// TwinCAT 3 PLC project AdsGo_Det
// Title: AdsClient_DeterministicTester
// Description: This project provides a series of programs and symbols to allow integration testing of ADS clients by utilising deterministic outputs on symbols based on writeable inputs (such as nSeed).
// ProgramVersion: 3.1.4026.25
// libraries:
//   Tc2_Standard, * (Beckhoff Automation GmbH)
//   Tc2_System, * (Beckhoff Automation GmbH)
//   Tc3_Module, * (Beckhoff Automation GmbH)
// project tree:
//   Lib/Arrays/ E_ArrayEnum.TcDUT, FB_ArrayTest.TcPOU, ST_Array.TcDUT, ST_ArrayBits.TcDUT
//   Lib/Attributes/ FB_AttributeTest.TcPOU
//   Lib/BitPacking/ FB_BitPackingTest.TcPOU, ST_BitPacking.TcDUT
//   Lib/Enums/ E_Int.TcDUT, E_Sparse.TcDUT, E_UInt.TcDUT, E_Default.TcDUT, E_Dint.TcDUT, E_Byte.TcDUT, E_Sint.TcDUT, E_USint.TcDUT, E_Word.TcDUT, E_ULint.TcDUT, E_UDint.TcDUT, E_Lint.TcDUT, E_DWord.TcDUT, E_LWord.TcDUT, E_Negative.TcDUT, FB_EnumTest.TcPOU
//   Lib/ FB_TickCounter.TcPOU
//   Lib/Gvl/ FB_GvlTest.TcPOU, GVL_Test.TcGVL
//   Lib/Strings/ FB_StringTest.TcPOU
//   Lib/StructPacking/ FB_StructPackingTest.TcPOU, ST_StructPackEight.TcDUT, ST_StructPackFour.TcDUT, ST_StructPackNone.TcDUT, ST_StructPackTwo.TcDUT
//   Lib/Types/ FB_TypeTest.TcPOU, ST_TypeTestStruct.TcDUT, ST_TypeTestSubStruct.TcDUT
//   Lib/Writing/ FB_WriteTest.TcPOU
//   Programs/ Main.TcPOU
//   Tasks/ PlcTask.TcTTO
// real-time tasks:
//   TASK PlcTask: cycle T#10ms, priority 20, ADS port 354

CONFIGURATION AdsGo_Det
    RESOURCE PLC ON TwinCAT3
        TASK PlcTask(INTERVAL := T#10ms, PRIORITY := 20);
        PROGRAM Main WITH PlcTask : Main;
    END_RESOURCE
END_CONFIGURATION

// ---- Lib/Arrays/E_ArrayEnum.TcDUT
{attribute 'qualified_only'}
{attribute 'strict'}
{attribute 'to_string'}
TYPE E_ArrayEnum :
(
	Member1 := 0,
	Member2,
	Member3,
	Member4
);
END_TYPE

// ---- Lib/Arrays/ST_Array.TcDUT
TYPE ST_Array :
STRUCT
	arr1 : ARRAY[0..2,0..2] OF INT;
	arr2 : ARRAY[0..1,0..1] OF ARRAY[0..1,0..1] OF INT;
	arr3 : ARRAY[0..1,0..1,0..1] OF ARRAY[0..1] OF INT;
END_STRUCT
END_TYPE

// ---- Lib/Arrays/ST_ArrayBits.TcDUT
TYPE ST_ArrayBits :
STRUCT
	bBit0 : BIT;
	bBit1 : BIT;
	bBit2 : BIT;
	bBit3 : BIT;
	bBit4 : BIT;
	bBit5 : BIT;
	bBit6 : BIT;
	bBit7 : BIT;
	bBit8 : BIT;
	bBit9 : BIT;
	bBit10 : BIT;
	bBit11 : BIT;
	bBit12 : BIT;
	bBit13 : BIT;
	bBit14 : BIT;
	bBit15 : BIT;
	bBit16 : BIT;
	bBit17 : BIT;
	bBit18 : BIT;
	bBit19 : BIT;
	bBit20 : BIT;
	bBit21 : BIT;
	bBit22 : BIT;
	bBit23 : BIT;
	bBit24 : BIT;
	bBit25 : BIT;
	bBit26 : BIT;
	bBit27 : BIT;
	bBit28 : BIT;
	bBit29 : BIT;
	bBit30 : BIT;
	bBit31 : BIT;
	bBit32 : BIT;
	bBit33 : BIT;
	bBit34 : BIT;
	bBit35 : BIT;
	bBit36 : BIT;
	bBit37 : BIT;
	bBit38 : BIT;
	bBit39 : BIT;
	bBit40 : BIT;
	bBit41 : BIT;
	bBit42 : BIT;
	bBit43 : BIT;
	bBit44 : BIT;
	bBit45 : BIT;
	bBit46 : BIT;
	bBit47 : BIT;
	bBit48 : BIT;
	bBit49 : BIT;
	bBit50 : BIT;
	bBit51 : BIT;
	bBit52 : BIT;
	bBit53 : BIT;
	bBit54 : BIT;
	bBit55 : BIT;
	bBit56 : BIT;
	bBit57 : BIT;
	bBit58 : BIT;
	bBit59 : BIT;
	bBit60 : BIT;
	bBit61 : BIT;
	bBit62 : BIT;
	bBit63 : BIT;
END_STRUCT
END_TYPE

// ---- Lib/BitPacking/ST_BitPacking.TcDUT
TYPE ST_BitPacking :
STRUCT
	bBit0 : BIT;
	bBit1 : BIT;
	bBit2 : BIT;
	bBit3 : BIT;
	bBit4 : BIT;
	bBit5 : BIT;
	bBit6 : BIT;
	bBit7 : BIT;
	bBit8 : BIT;
	bBit9 : BIT;
	bBit10 : BIT;
	bBit11 : BIT;
	bBit12 : BIT;
	bBit13 : BIT;
	bBit14 : BIT;
	bBit15 : BIT;
	bBit16 : BIT;
	bBit17 : BIT;
	bBit18 : BIT;
	bBit19 : BIT;
	bBit20 : BIT;
	bBit21 : BIT;
	bBit22 : BIT;
	bBit23 : BIT;
	bBit24 : BIT;
	bBit25 : BIT;
	bBit26 : BIT;
	bBit27 : BIT;
	bBit28 : BIT;
	bBit29 : BIT;
	bBit30 : BIT;
	bBit31 : BIT;
	bBit32 : BIT;
	bBit33 : BIT;
	bBit34 : BIT;
	bBit35 : BIT;
	bBit36 : BIT;
	bBit37 : BIT;
	bBit38 : BIT;
	bBit39 : BIT;
	bBit40 : BIT;
	bBit41 : BIT;
	bBit42 : BIT;
	bBit43 : BIT;
	bBit44 : BIT;
	bBit45 : BIT;
	bBit46 : BIT;
	bBit47 : BIT;
	bBit48 : BIT;
	bBit49 : BIT;
	bBit50 : BIT;
	bBit51 : BIT;
	bBit52 : BIT;
	bBit53 : BIT;
	bBit54 : BIT;
	bBit55 : BIT;
	bBit56 : BIT;
	bBit57 : BIT;
	bBit58 : BIT;
	bBit59 : BIT;
	bBit60 : BIT;
	bBit61 : BIT;
	bBit62 : BIT;
	bBit63 : BIT;
END_STRUCT
END_TYPE

// ---- Lib/Enums/E_Int.TcDUT
{attribute 'qualified_only'}
{attribute 'strict'}
{attribute 'to_string'}
TYPE E_Int :
(
	eOptionA := 0,
	eOptionB,
	eOptionC
) INT;
END_TYPE

// ---- Lib/Enums/E_Sparse.TcDUT
{attribute 'qualified_only'}
{attribute 'strict'}
{attribute 'to_string'}
TYPE E_Sparse :
(
	eOptionA := -10,
	eOptionB := 0,
	eOptionC := 100
);
END_TYPE

// ---- Lib/Enums/E_UInt.TcDUT
{attribute 'qualified_only'}
{attribute 'strict'}
{attribute 'to_string'}
TYPE E_UInt :
(
	eOptionA := 0,
	eOptionB,
	eOptionC
) UINT;
END_TYPE

// ---- Lib/Enums/E_Default.TcDUT
{attribute 'qualified_only'}
{attribute 'strict'}
{attribute 'to_string'}
TYPE E_Default :
(
	eOptionA := 0,
	eOptionB,
	eOptionC
);
END_TYPE

// ---- Lib/Enums/E_Dint.TcDUT
{attribute 'qualified_only'}
{attribute 'strict'}
{attribute 'to_string'}
TYPE E_Dint :
(
	eOptionA := 0,
	eOptionB,
	eOptionC
) DINT;
END_TYPE

// ---- Lib/Enums/E_Byte.TcDUT
{attribute 'qualified_only'}
{attribute 'strict'}
{attribute 'to_string'}
TYPE E_Byte :
(
	eOptionA := 0,
	eOptionB,
	eOptionC
) BYTE;
END_TYPE

// ---- Lib/Enums/E_Sint.TcDUT
{attribute 'qualified_only'}
{attribute 'strict'}
{attribute 'to_string'}
TYPE E_Sint :
(
	eOptionA := 0,
	eOptionB,
	eOptionC
) SINT;
END_TYPE

// ---- Lib/Enums/E_USint.TcDUT
{attribute 'qualified_only'}
{attribute 'strict'}
{attribute 'to_string'}
TYPE E_USint :
(
	eOptionA := 0,
	eOptionB,
	eOptionC
) USINT;
END_TYPE

// ---- Lib/Enums/E_Word.TcDUT
{attribute 'qualified_only'}
{attribute 'strict'}
{attribute 'to_string'}
TYPE E_Word :
(
	eOptionA := 0,
	eOptionB,
	eOptionC
) WORD;
END_TYPE

// ---- Lib/Enums/E_ULint.TcDUT
{attribute 'qualified_only'}
{attribute 'strict'}
{attribute 'to_string'}
TYPE E_ULint :
(
	eOptionA := 0,
	eOptionB,
	eOptionC
) ULINT;
END_TYPE

// ---- Lib/Enums/E_UDint.TcDUT
{attribute 'qualified_only'}
{attribute 'strict'}
{attribute 'to_string'}
TYPE E_UDint :
(
	eOptionA := 0,
	eOptionB,
	eOptionC
) UDINT;
END_TYPE

// ---- Lib/Enums/E_Lint.TcDUT
{attribute 'qualified_only'}
{attribute 'strict'}
{attribute 'to_string'}
TYPE E_Lint :
(
	eOptionA := 0,
	eOptionB,
	eOptionC
) LINT;
END_TYPE

// ---- Lib/Enums/E_DWord.TcDUT
{attribute 'qualified_only'}
{attribute 'strict'}
{attribute 'to_string'}
TYPE E_DWord :
(
	eOptionA := 0,
	eOptionB,
	eOptionC
) DWORD;
END_TYPE

// ---- Lib/Enums/E_LWord.TcDUT
{attribute 'qualified_only'}
{attribute 'strict'}
{attribute 'to_string'}
TYPE E_LWord :
(
	eOptionA := 0,
	eOptionB,
	eOptionC
) LWORD;
END_TYPE

// ---- Lib/Enums/E_Negative.TcDUT
{attribute 'qualified_only'}
{attribute 'strict'}
{attribute 'to_string'}
TYPE E_Negative :
(
	eOptionA := -1,
	eOptionB := 0,
	eOptionC := 1
);
END_TYPE

// ---- Lib/StructPacking/ST_StructPackEight.TcDUT
{attribute 'pack_mode' := '8'}
TYPE ST_StructPackEight :
STRUCT
	bBoolMember1 : BOOL;
	nDwordMember : DWORD;
	bBoolMember2 : BOOL;
	nLwordMember : LWORD;
END_STRUCT
END_TYPE

// ---- Lib/StructPacking/ST_StructPackFour.TcDUT
{attribute 'pack_mode' := '4'}
TYPE ST_StructPackFour :
STRUCT
	bBoolMember1 : BOOL;
	nDwordMember : DWORD;
	bBoolMember2 : BOOL;
	nLwordMember : LWORD;
END_STRUCT
END_TYPE

// ---- Lib/StructPacking/ST_StructPackNone.TcDUT
{attribute 'pack_mode' := '0'}
TYPE ST_StructPackNone :
STRUCT
	bBoolMember1 : BOOL;
	nDwordMember : DWORD;
	bBoolMember2 : BOOL;
	nLwordMember : LWORD;
END_STRUCT
END_TYPE

// ---- Lib/StructPacking/ST_StructPackTwo.TcDUT
{attribute 'pack_mode' := '2'}
TYPE ST_StructPackTwo :
STRUCT
	bBoolMember1 : BOOL;
	nDwordMember : DWORD;
	bBoolMember2 : BOOL;
	nLwordMember : LWORD;
END_STRUCT
END_TYPE

// ---- Lib/Types/ST_TypeTestStruct.TcDUT
TYPE ST_TypeTestStruct :
STRUCT
	// Control (writable by Go test)
	nSeed : UDINT := 0;
	bAutoMode : BOOL := FALSE;
	nAutoTickInterval : UDINT := 50;

	// Outputs
	bBoolVar : BOOL;
	nSintVar : SINT;
	nUsintVar : USINT;
	nByteVar : BYTE;
	nIntVar : INT;
	nUintVar : UINT;
	nWordVar : WORD;
	nDintVar : DINT;
	nUdintVar : UDINT;
	nDwordVar : DWORD;
	nLintVar : LINT;
	nUlintVar : ULINT;
	nLwordVar : LWORD;
	fRealVar : REAL;
	fLrealVar : LREAL;
	tTimeVar : TIME;
	tdTimeOfDayVar : TOD;
	dDateVar : DATE;
	dtDateTimeVar : DT;
	tLtimeVar : LTIME;
	tdLTimeOfDayVar : LTOD;
	dLDateVar : LDATE;
	dtLDateTimeVar : LDT;
	sStringVar : STRING(255);
	stSubStructVar : ST_TypeTestSubStruct;
END_STRUCT
END_TYPE

// ---- Lib/Types/ST_TypeTestSubStruct.TcDUT
TYPE ST_TypeTestSubStruct :
STRUCT
	// Outputs
	bBoolVar : BOOL;
	nSintVar : SINT;
	nUsintVar : USINT;
	nByteVar : BYTE;
	nIntVar : INT;
	nUintVar : UINT;
	nWordVar : WORD;
	nDintVar : DINT;
	nUdintVar : UDINT;
	nDwordVar : DWORD;
	nLintVar : LINT;
	nUlintVar : ULINT;
	nLwordVar : LWORD;
	fRealVar : REAL;
	fLrealVar : LREAL;
	tTimeVar : TIME;
	tdTimeOfDayVar : TOD;
	dDateVar : DATE;
	dtDateTimeVar : DT;
	tLtimeVar : LTIME;
	tdLTimeOfDayVar : LTOD;
	dLDateVar : LDATE;
	dtLDateTimeVar : LDT;
	sStringVar : STRING(255);
END_STRUCT
END_TYPE

// ---- Lib/Gvl/GVL_Test.TcGVL
{attribute 'qualified_only'}
VAR_GLOBAL
	bBoolVar : BOOL;
	nSintVar : SINT;
	nUsintVar : USINT;
	nByteVar : BYTE;
	nIntVar : INT;
	nUintVar : UINT;
	nWordVar : WORD;
	nDintVar : DINT;
	nUdintVar : UDINT;
	nDwordVar : DWORD;
	nLintVar : LINT;
	nUlintVar : ULINT;
	nLwordVar : LWORD;
	fRealVar : REAL;
	fLrealVar : LREAL;
	tTimeVar : TIME;
	tdTimeOfDayVar : TOD;
	dDateVar : DATE;
	dtDateTimeVar : DT;
	tLtimeVar : LTIME;
	tdLTimeOfDayVar : LTOD;
	dLDateVar : LDATE;
	dtLDateTimeVar : LDT;
	sStringVar : STRING(255);
	stStructVar : ST_TypeTestStruct;
	aIntArray : ARRAY[0..9] OF INT;
	aDintArray : ARRAY[0..9] OF DINT;
	aIntArray2d : ARRAY[0..2, 0..2] OF INT;
END_VAR

// ---- Programs/Main.TcPOU
PROGRAM Main
VAR
	nSeed : ULINT := 0;
	fbTickCounter : FB_TickCounter;
	bAutoMode : BOOL := FALSE;
	nAutoTickInterval : UDINT := 50;
	
	fbTypeTest : FB_TypeTest(nSeed := nSeed);
	fbStringTest : FB_StringTest(nSeed := nSeed);
	fbStructTest : FB_StructPackingTest(nSeed := nSeed);
	fbEnumTest : FB_EnumTest(nSeed := nSeed);
	fbBitPackingTest : FB_BitPackingTest(nSeed := nSeed);
	fbArrayTest : FB_ArrayTest(nSeed := nSeed);
	fbWriteTest : FB_WriteTest;
	
	fbGvlTest : FB_GvlTest(nSeed := nSeed);
	
	{attribute 'some_made_up_var_key':='some_made_up_var_value'}
	fbAttributeTest : FB_AttributeTest;	
END_VAR

fbTypeTest();
fbStringTest();
fbStructTest();
fbEnumTest();
fbBitPackingTest();
fbArrayTest();
fbWriteTest();

fbGvlTest();

fbAttributeTest();

fbTickCounter(bExecute := bAutoMode, nAutoTickInterval := nAutoTickInterval);

IF bAutoMode AND fbTickCounter.bTrigger THEN
	nSeed := nSeed + 1;
END_IF

END_PROGRAM

// ---- Lib/FB_TickCounter.TcPOU
FUNCTION_BLOCK FB_TickCounter
VAR_INPUT
	bExecute : BOOL := FALSE;
	nAutoTickInterval : UDINT := 50;
END_VAR
VAR_OUTPUT
	bTrigger : BOOL;
END_VAR
VAR
	nSeed : REFERENCE TO UDINT;
	nTickCounter : UDINT;
END_VAR

bTrigger := bExecute AND nTickCounter >= nAutoTickInterval;

IF bExecute THEN
	IF bTrigger THEN
		nTickCounter := 0;
	ELSE
		nTickCounter := nTickCounter + 1;
	END_IF
ELSE
	nTickCounter := 0;
END_IF

END_FUNCTION_BLOCK

// ---- Lib/Types/FB_TypeTest.TcPOU
FUNCTION_BLOCK FB_TypeTest
VAR
	// Control
	nSeed : REFERENCE TO ULINT;

	// Outputs
	bBoolVar : BOOL;
	nSintVar : SINT;
	nUsintVar : USINT;
	nByteVar : BYTE;
	nIntVar : INT;
	nUintVar : UINT;
	nWordVar : WORD;
	nDintVar : DINT;
	nUdintVar : UDINT;
	nDwordVar : DWORD;
	nLintVar : LINT;
	nUlintVar : ULINT;
	nLwordVar : LWORD;
	fRealVar : REAL;
	fLrealVar : LREAL;
	
	nSubRange : INT(-10..10);
	
	tTimeVar : TIME;
	tdTimeOfDayVar : TOD;
	dDateVar : DATE;
	dtDateTimeVar : DT;
	tLtimeVar : LTIME;
	tdLTimeOfDayVar : LTOD;
	dLDateVar : LDATE;
	dtLDateTimeVar : LDT;
	
	sStringVar : STRING(255);
	stStructVar : ST_TypeTestStruct;
	
	aIntArray : ARRAY[0..9] OF INT;
	aDintArray : ARRAY[-9..9] OF DINT;
	aIntArray2d : ARRAY[0..2, 0..2] OF INT;
	aStructVar : ARRAY[0..9] OF ST_TypeTestSubStruct;

	// Private
	nLoopIndex1 : DINT;
	nLoopIndex2 : UDINT;
END_VAR

// -----------------------------------------------------------------------
// Update variables — all fields are deterministic functions of seed
// -----------------------------------------------------------------------
bBoolVar := (nSeed MOD 2 = 0);
nSintVar := ULINT_TO_SINT(nSeed);
nUsintVar := ULINT_TO_USINT(nSeed);
nByteVar := ULINT_TO_BYTE(nSeed);
nIntVar := ULINT_TO_INT(nSeed);
nUintVar := ULINT_TO_UINT(nSeed);
nWordVar := ULINT_TO_WORD(nSeed);
nDintVar := ULINT_TO_DINT(nSeed);
nUdintVar := ULINT_TO_UDINT(nSeed);
nDwordVar := ULINT_TO_DWORD(nSeed);
nLintVar := ULINT_TO_LINT(nSeed);
nUlintVar := nSeed;
nLwordVar := ULINT_TO_LWORD(nSeed);
fRealVar := ULINT_TO_REAL(nSeed);
fLrealVar := ULINT_TO_LREAL(nSeed);

// Sub range
nSubRange := ULINT_TO_INT(nSeed MOD 21) - 10;

// Date/time types — raw truncating casts, same bit pattern Go test will verify
tTimeVar := ULINT_TO_TIME(nSeed);
tdTimeOfDayVar := ULINT_TO_TOD(nSeed MOD 86400000);
dDateVar := ULINT_TO_DATE(nSeed);
dtDateTimeVar := ULINT_TO_DT(nSeed);
tLTimeVar := ULINT_TO_LTIME(nSeed);
tdLTimeOfDayVar  := ULINT_TO_LTOD(nSeed MOD 86400000000000);
dLDateVar := ULINT_TO_LDATE(nSeed);
dtLDateTimeVar := ULINT_TO_LDT(nSeed);
sStringVar := CONCAT('S=', ULINT_TO_STRING(nSeed));

// -----------------------------------------------------------------------
// Update test struct — all fields are deterministic functions of seed
// -----------------------------------------------------------------------
stStructVar.nSeed := ULINT_TO_UDINT(nSeed);

stStructVar.bBoolVar := bBoolVar;
stStructVar.nSintVar := nSintVar;
stStructVar.nUsintVar := nUsintVar;
stStructVar.nByteVar := nByteVar;
stStructVar.nIntVar := nIntVar;
stStructVar.nUintVar := nUintVar;
stStructVar.nWordVar := nWordVar;
stStructVar.nDintVar := nDintVar;
stStructVar.nUdintVar := nUdintVar;
stStructVar.nDwordVar := nDwordVar;
stStructVar.nLintVar := nLintVar;
stStructVar.nUlintVar := nUlintVar;
stStructVar.nLwordVar := nLwordVar;
stStructVar.fRealVar := fRealVar;
stStructVar.fLrealVar := fLrealVar;
stStructVar.tTimeVar := tTimeVar;
stStructVar.tdTimeOfDayVar := tdTimeOfDayVar;
stStructVar.dDateVar := dDateVar;
stStructVar.dtDateTimeVar := dtDateTimeVar;
stStructVar.tLTimeVar := tLTimeVar;
stStructVar.tdLTimeOfDayVar := tdLTimeOfDayVar;
stStructVar.dLDateVar := dLDateVar;
stStructVar.dtLDateTimeVar := dtLDateTimeVar;
stStructVar.sStringVar := sStringVar;

// Nested struct
stStructVar.stSubStructVar.bBoolVar := bBoolVar;
stStructVar.stSubStructVar.nSintVar := nSintVar;
stStructVar.stSubStructVar.nUsintVar := nUsintVar;
stStructVar.stSubStructVar.nByteVar := nByteVar;
stStructVar.stSubStructVar.nIntVar := nIntVar;
stStructVar.stSubStructVar.nUintVar := nUintVar;
stStructVar.stSubStructVar.nWordVar := nWordVar;
stStructVar.stSubStructVar.nDintVar := nDintVar;
stStructVar.stSubStructVar.nUdintVar := nUdintVar;
stStructVar.stSubStructVar.nDwordVar := nDwordVar;
stStructVar.stSubStructVar.nLintVar := nLintVar;
stStructVar.stSubStructVar.nUlintVar := nUlintVar;
stStructVar.stSubStructVar.nLwordVar := nLwordVar;
stStructVar.stSubStructVar.fRealVar := fRealVar;
stStructVar.stSubStructVar.fLrealVar := fLrealVar;
stStructVar.stSubStructVar.tTimeVar := tTimeVar;
stStructVar.stSubStructVar.tdTimeOfDayVar := tdTimeOfDayVar;
stStructVar.stSubStructVar.dDateVar := dDateVar;
stStructVar.stSubStructVar.dtDateTimeVar := dtDateTimeVar;
stStructVar.stSubStructVar.tLTimeVar := tLTimeVar;
stStructVar.stSubStructVar.tdLTimeOfDayVar := tdLTimeOfDayVar;
stStructVar.stSubStructVar.dLDateVar := dLDateVar;
stStructVar.stSubStructVar.dtLDateTimeVar := dtLDateTimeVar;
stStructVar.stSubStructVar.sStringVar := sStringVar;

// -----------------------------------------------------------------------
// Update 1-D arrays: element[i] = UDINT_TO_x(seed + i)
// -----------------------------------------------------------------------
FOR nLoopIndex1 := 0 TO 9 DO
	aIntArray[nLoopIndex1] := ULINT_TO_INT(nSeed + DINT_TO_ULINT(nLoopIndex1));
END_FOR

FOR nLoopIndex1 := -9 TO 9 DO
	aDintArray[nLoopIndex1] := ULINT_TO_DINT(nSeed) + nLoopIndex1;
END_FOR

// -----------------------------------------------------------------------
// Update 2-D array: element[i,j] = UDINT_TO_INT(seed + i*3 + j)
// -----------------------------------------------------------------------
FOR nLoopIndex1 := 0 TO 2 DO
	FOR nLoopIndex2 := 0 TO 2 DO
		aIntArray2d[nLoopIndex1, nLoopIndex2] := LINT_TO_INT(ULINT_TO_LINT(nSeed) + nLoopIndex1 * 3 + nLoopIndex2);
	END_FOR
END_FOR

// -----------------------------------------------------------------------
// Update struct array: 
// -----------------------------------------------------------------------
FOR nLoopIndex1 := 0 TO 9 DO
	aStructVar[nLoopIndex1].bBoolVar := bBoolVar;
	aStructVar[nLoopIndex1].nSintVar := nSintVar;
	aStructVar[nLoopIndex1].nUsintVar := nUsintVar;
	aStructVar[nLoopIndex1].nByteVar := nByteVar;
	aStructVar[nLoopIndex1].nIntVar := nIntVar;
	aStructVar[nLoopIndex1].nUintVar := nUintVar;
	aStructVar[nLoopIndex1].nWordVar := nWordVar;
	aStructVar[nLoopIndex1].nDintVar := nDintVar;
	aStructVar[nLoopIndex1].nUdintVar := nUdintVar;
	aStructVar[nLoopIndex1].nDwordVar := nDwordVar;
	aStructVar[nLoopIndex1].nLintVar := nLintVar;
	aStructVar[nLoopIndex1].nUlintVar := nUlintVar;
	aStructVar[nLoopIndex1].nLwordVar := nLwordVar;
	aStructVar[nLoopIndex1].fRealVar := fRealVar;
	aStructVar[nLoopIndex1].fLrealVar := fLrealVar;
	aStructVar[nLoopIndex1].tTimeVar := tTimeVar;
	aStructVar[nLoopIndex1].tdTimeOfDayVar := tdTimeOfDayVar;
	aStructVar[nLoopIndex1].dDateVar := dDateVar;
	aStructVar[nLoopIndex1].dtDateTimeVar := dtDateTimeVar;
	aStructVar[nLoopIndex1].tLTimeVar := tLTimeVar;
	aStructVar[nLoopIndex1].tdLTimeOfDayVar := tdLTimeOfDayVar;
	aStructVar[nLoopIndex1].dLDateVar := dLDateVar;
	aStructVar[nLoopIndex1].dtLDateTimeVar := dtLDateTimeVar;
	aStructVar[nLoopIndex1].sStringVar := sStringVar;
END_FOR

//FB_Init is always available implicitly and it is used primarily for initialization.
//The return value is not evaluated. For a specific influence, you can also declare the
//methods explicitly and provide additional code there with the standard initialization
//code. You can evaluate the return value.
METHOD FB_Init: BOOL
VAR_INPUT
    bInitRetains : BOOL; // TRUE: the retain variables are initialized (reset warm / reset cold)
    bInCopyCode : BOOL;  // TRUE: the instance will be copied to the copy code afterward (online change)
	nSeed : REFERENCE TO ULINT;
END_VAR
THIS^.nSeed REF= nSeed;
END_METHOD

END_FUNCTION_BLOCK

// ---- Lib/Strings/FB_StringTest.TcPOU
FUNCTION_BLOCK FB_StringTest
VAR
	// Control
	nSeed : REFERENCE TO ULINT;

	// Written by the Go test
	sStringVar : STRING(255);
	sShortStringVar : STRING(5);
	wsWStringVar : WSTRING(255);

	// What the PLC sees in them, recomputed every cycle
	nStringLen : INT;                        // LEN(sStringVar): characters as the PLC counts them
	nShortStringLen : INT;                   // LEN(sShortStringVar)
	nWStringLen : INT;                       // WLEN(wsWStringVar): UTF-16 code units
	aStringBytes : ARRAY[0..255] OF BYTE;    // the bytes of sStringVar
	aWStringWords : ARRAY[0..255] OF WORD;   // the code units of wsWStringVar
	wsFromString : WSTRING(255);             // STRING_TO_WSTRING(sStringVar)
	sFromWString : STRING(255);              // WSTRING_TO_STRING(wsWStringVar)

	// Produced by the PLC
	sLatinLiteral : STRING(255) := 'Grüße € ÄÖÜ ñ ©';
	wsLiteral : WSTRING(255) := "Grüße € 日本語";
	sAllBytes : STRING(255);                 // bytes 16#01..16#FF in order
	wsAllBytes : WSTRING(255);               // STRING_TO_WSTRING(sAllBytes): Beckhoff's mapping of every byte

	// Private
	aByteTable : ARRAY[0..255] OF BYTE;
	nIndex : INT;
END_VAR

// -----------------------------------------------------------------------
// Report what the PLC sees in the strings the Go test wrote
// -----------------------------------------------------------------------
nStringLen := LEN(sStringVar);
nShortStringLen := LEN(sShortStringVar);
nWStringLen := WLEN(wsWStringVar);
MEMCPY(destAddr := ADR(aStringBytes), srcAddr := ADR(sStringVar), n := SIZEOF(aStringBytes));
MEMCPY(destAddr := ADR(aWStringWords), srcAddr := ADR(wsWStringVar), n := SIZEOF(aWStringWords));
wsFromString := STRING_TO_WSTRING(sStringVar);
sFromWString := WSTRING_TO_STRING(wsWStringVar);

// -----------------------------------------------------------------------
// Every non-NUL byte in one STRING, and Beckhoff's conversion of it
// -----------------------------------------------------------------------
FOR nIndex := 0 TO 254 DO
	aByteTable[nIndex] := INT_TO_BYTE(nIndex + 1);
END_FOR
aByteTable[255] := 0;
MEMCPY(destAddr := ADR(sAllBytes), srcAddr := ADR(aByteTable), n := SIZEOF(sAllBytes));
wsAllBytes := STRING_TO_WSTRING(sAllBytes);

//FB_Init is always available implicitly and it is used primarily for initialization.
//The return value is not evaluated. For a specific influence, you can also declare the
//methods explicitly and provide additional code there with the standard initialization
//code. You can evaluate the return value.
METHOD FB_Init: BOOL
VAR_INPUT
    bInitRetains : BOOL; // TRUE: the retain variables are initialized (reset warm / reset cold)
    bInCopyCode : BOOL;  // TRUE: the instance will be copied to the copy code afterward (online change)
	nSeed : REFERENCE TO ULINT;
END_VAR
THIS^.nSeed REF= nSeed;
END_METHOD

END_FUNCTION_BLOCK

// ---- Lib/StructPacking/FB_StructPackingTest.TcPOU
{attribute 'linkalways'}
FUNCTION_BLOCK FB_StructPackingTest
VAR
	nSeed : REFERENCE TO ULINT;
	stPackNone : ST_StructPackNone;
	stPackTwo : ST_StructPackTwo;
	stPackFour : ST_StructPackFour;
	stPackEight : ST_StructPackEight;
	
	// pack_*_write: Go-owned write targets (PLC never modifies, used in phase 2)
	stPackNoneWrite : ST_StructPackNone;
	stPackTwoWrite : ST_StructPackTwo;
	stPackFourWrite : ST_StructPackFour;
	stPackEightWrite : ST_StructPackEight;
END_VAR

// All four structs share the same fields and the same seed-driven formula.
// b1  = (seed MOD 2 = 0)
// d1  = seed
// b2  = (seed MOD 3 = 0)
// lw1 = LWORD(seed) * LWORD(3)
stPackNone.bBoolMember1 := (nSeed MOD 2 = 0);
stPackNone.nDwordMember := ULINT_TO_DWORD(nSeed);
stPackNone.bBoolMember2 := (nSeed MOD 3 = 0);
stPackNone.nLwordMember := ULINT_TO_LWORD(nSeed) * UDINT_TO_LWORD(3);

stPackTwo.bBoolMember1 := stPackNone.bBoolMember1;
stPackTwo.nDwordMember := stPackNone.nDwordMember;
stPackTwo.bBoolMember2 := stPackNone.bBoolMember2;
stPackTwo.nLwordMember := stPackNone.nLwordMember;

stPackFour.bBoolMember1 := stPackNone.bBoolMember1;
stPackFour.nDwordMember := stPackNone.nDwordMember;
stPackFour.bBoolMember2 := stPackNone.bBoolMember2;
stPackFour.nLwordMember := stPackNone.nLwordMember;

stPackEight.bBoolMember1 := stPackNone.bBoolMember1;
stPackEight.nDwordMember := stPackNone.nDwordMember;
stPackEight.bBoolMember2 := stPackNone.bBoolMember2;
stPackEight.nLwordMember := stPackNone.nLwordMember;

//FB_Init is always available implicitly and it is used primarily for initialization.
//The return value is not evaluated. For a specific influence, you can also declare the
//methods explicitly and provide additional code there with the standard initialization
//code. You can evaluate the return value.
METHOD FB_Init: BOOL
VAR_INPUT
    bInitRetains : BOOL; // TRUE: the retain variables are initialized (reset warm / reset cold)
    bInCopyCode : BOOL;  // TRUE: the instance will be copied to the copy code afterward (online change)
	nSeed : REFERENCE TO ULINT;
END_VAR
THIS^.nSeed REF= nSeed;
END_METHOD

END_FUNCTION_BLOCK

// ---- Lib/Enums/FB_EnumTest.TcPOU
FUNCTION_BLOCK FB_EnumTest
VAR
	// Control
	nSeed : REFERENCE TO ULINT;

	// Outputs
	eDefault : E_Default;
	eByte : E_Byte;
	eWord : E_Word;
	eDWord : E_DWord;
	eLWord : E_LWord;
	eSInt : E_SInt;
	eUSInt : E_USInt;
	eInt : E_Int;
	eUInt : E_UInt;
	eDInt : E_DInt;
	eUDInt : E_UDInt;
	eLInt : E_LInt;
	eULInt : E_ULInt;
	eNegative : E_Negative;
	eSparse : E_Sparse;
	
	eDefaultWrite : E_Default;
	eByteWrite : E_Byte;
	eWordWrite : E_Word;
	eDWordWrite : E_DWord;
	eLWordWrite : E_LWord;
	eSIntWrite : E_SInt;
	eUSIntWrite : E_USInt;
	eIntWrite : E_Int;
	eUIntWrite : E_UInt;
	eDIntWrite : E_DInt;
	eUDIntWrite : E_UDInt;
	eLIntWrite : E_LInt;
	eULIntWrite : E_ULInt;
	eNegativeWrite : E_Negative;
	eSparseWrite : E_Sparse;
	
	eImplicit : (eImplicitOptionA, eImplicitOptionB, eImplicitOptionC);
END_VAR

CASE nSeed MOD 3 OF
	0: eDefault := E_Default.eOptionA;
	1: eDefault := E_Default.eOptionB;
	2: eDefault := E_Default.eOptionC;
END_CASE

// BYTE
CASE eDefault OF
	E_Default.eOptionA: eByte := E_Byte.eOptionA;
	E_Default.eOptionB: eByte := E_Byte.eOptionB;
	E_Default.eOptionC: eByte := E_Byte.eOptionC;
END_CASE

// WORD
CASE eDefault OF
	E_Default.eOptionA: eWord := E_Word.eOptionA;
	E_Default.eOptionB: eWord := E_Word.eOptionB;
	E_Default.eOptionC: eWord := E_Word.eOptionC;
END_CASE

// DWORD
CASE eDefault OF
	E_Default.eOptionA: eDWord := E_DWord.eOptionA;
	E_Default.eOptionB: eDWord := E_DWord.eOptionB;
	E_Default.eOptionC: eDWord := E_DWord.eOptionC;
END_CASE

// LWORD
CASE eDefault OF
	E_Default.eOptionA: eLWord := E_LWord.eOptionA;
	E_Default.eOptionB: eLWord := E_LWord.eOptionB;
	E_Default.eOptionC: eLWord := E_LWord.eOptionC;
END_CASE

// SINT
CASE eDefault OF
	E_Default.eOptionA: eSInt := E_SInt.eOptionA;
	E_Default.eOptionB: eSInt := E_SInt.eOptionB;
	E_Default.eOptionC: eSInt := E_SInt.eOptionC;
END_CASE

// USINT
CASE eDefault OF
	E_Default.eOptionA: eUSInt := E_USInt.eOptionA;
	E_Default.eOptionB: eUSInt := E_USInt.eOptionB;
	E_Default.eOptionC: eUSInt := E_USInt.eOptionC;
END_CASE

// INT
CASE eDefault OF
	E_Default.eOptionA: eInt := E_Int.eOptionA;
	E_Default.eOptionB: eInt := E_Int.eOptionB;
	E_Default.eOptionC: eInt := E_Int.eOptionC;
END_CASE

// UINT
CASE eDefault OF
	E_Default.eOptionA: eUInt := E_UInt.eOptionA;
	E_Default.eOptionB: eUInt := E_UInt.eOptionB;
	E_Default.eOptionC: eUInt := E_UInt.eOptionC;
END_CASE

// DINT
CASE eDefault OF
	E_Default.eOptionA: eDInt := E_DInt.eOptionA;
	E_Default.eOptionB: eDInt := E_DInt.eOptionB;
	E_Default.eOptionC: eDInt := E_DInt.eOptionC;
END_CASE

// UDINT
CASE eDefault OF
	E_Default.eOptionA: eUDInt := E_UDInt.eOptionA;
	E_Default.eOptionB: eUDInt := E_UDInt.eOptionB;
	E_Default.eOptionC: eUDInt := E_UDInt.eOptionC;
END_CASE

// LINT
CASE eDefault OF
	E_Default.eOptionA: eLInt := E_LInt.eOptionA;
	E_Default.eOptionB: eLInt := E_LInt.eOptionB;
	E_Default.eOptionC: eLInt := E_LInt.eOptionC;
END_CASE

// ULINT
CASE eDefault OF
	E_Default.eOptionA: eULInt := E_ULInt.eOptionA;
	E_Default.eOptionB: eULInt := E_ULInt.eOptionB;
	E_Default.eOptionC: eULInt := E_ULInt.eOptionC;
END_CASE

// Negative
CASE eDefault OF
	E_Default.eOptionA: eNegative := E_Negative.eOptionA;
	E_Default.eOptionB: eNegative := E_Negative.eOptionB;
	E_Default.eOptionC: eNegative := E_Negative.eOptionC;
END_CASE

// Sparse
CASE eDefault OF
	E_Default.eOptionA: eSparse := E_Sparse.eOptionA;
	E_Default.eOptionB: eSparse := E_Sparse.eOptionB;
	E_Default.eOptionC: eSparse := E_Sparse.eOptionC;
END_CASE

// Implicit
CASE eDefault OF
	E_Default.eOptionA: eImplicit := eImplicitOptionA;
	E_Default.eOptionB: eImplicit := eImplicitOptionB;
	E_Default.eOptionC: eImplicit := eImplicitOptionC;
END_CASE

//FB_Init is always available implicitly and it is used primarily for initialization.
//The return value is not evaluated. For a specific influence, you can also declare the
//methods explicitly and provide additional code there with the standard initialization
//code. You can evaluate the return value.
METHOD FB_Init: BOOL
VAR_INPUT
    bInitRetains : BOOL; // TRUE: the retain variables are initialized (reset warm / reset cold)
    bInCopyCode : BOOL;  // TRUE: the instance will be copied to the copy code afterward (online change)
	nSeed : REFERENCE TO ULINT;
END_VAR
THIS^.nSeed REF= nSeed;
END_METHOD

END_FUNCTION_BLOCK

// ---- Lib/BitPacking/FB_BitPackingTest.TcPOU
FUNCTION_BLOCK FB_BitPackingTest
VAR
	// Control
	nSeed : REFERENCE TO ULINT;

	// Outputs: bBitN = bit N of nSeed
	stBitPacking : ST_BitPacking;

	// Go-owned write target: the PLC never touches it
	stBitPackingWrite : ST_BitPacking;
END_VAR

// -----------------------------------------------------------------------
// bBitN := bit N of nSeed
// -----------------------------------------------------------------------
stBitPacking.bBit0 := (SHR(nSeed, 0) AND 1) = 1;
stBitPacking.bBit1 := (SHR(nSeed, 1) AND 1) = 1;
stBitPacking.bBit2 := (SHR(nSeed, 2) AND 1) = 1;
stBitPacking.bBit3 := (SHR(nSeed, 3) AND 1) = 1;
stBitPacking.bBit4 := (SHR(nSeed, 4) AND 1) = 1;
stBitPacking.bBit5 := (SHR(nSeed, 5) AND 1) = 1;
stBitPacking.bBit6 := (SHR(nSeed, 6) AND 1) = 1;
stBitPacking.bBit7 := (SHR(nSeed, 7) AND 1) = 1;
stBitPacking.bBit8 := (SHR(nSeed, 8) AND 1) = 1;
stBitPacking.bBit9 := (SHR(nSeed, 9) AND 1) = 1;
stBitPacking.bBit10 := (SHR(nSeed, 10) AND 1) = 1;
stBitPacking.bBit11 := (SHR(nSeed, 11) AND 1) = 1;
stBitPacking.bBit12 := (SHR(nSeed, 12) AND 1) = 1;
stBitPacking.bBit13 := (SHR(nSeed, 13) AND 1) = 1;
stBitPacking.bBit14 := (SHR(nSeed, 14) AND 1) = 1;
stBitPacking.bBit15 := (SHR(nSeed, 15) AND 1) = 1;
stBitPacking.bBit16 := (SHR(nSeed, 16) AND 1) = 1;
stBitPacking.bBit17 := (SHR(nSeed, 17) AND 1) = 1;
stBitPacking.bBit18 := (SHR(nSeed, 18) AND 1) = 1;
stBitPacking.bBit19 := (SHR(nSeed, 19) AND 1) = 1;
stBitPacking.bBit20 := (SHR(nSeed, 20) AND 1) = 1;
stBitPacking.bBit21 := (SHR(nSeed, 21) AND 1) = 1;
stBitPacking.bBit22 := (SHR(nSeed, 22) AND 1) = 1;
stBitPacking.bBit23 := (SHR(nSeed, 23) AND 1) = 1;
stBitPacking.bBit24 := (SHR(nSeed, 24) AND 1) = 1;
stBitPacking.bBit25 := (SHR(nSeed, 25) AND 1) = 1;
stBitPacking.bBit26 := (SHR(nSeed, 26) AND 1) = 1;
stBitPacking.bBit27 := (SHR(nSeed, 27) AND 1) = 1;
stBitPacking.bBit28 := (SHR(nSeed, 28) AND 1) = 1;
stBitPacking.bBit29 := (SHR(nSeed, 29) AND 1) = 1;
stBitPacking.bBit30 := (SHR(nSeed, 30) AND 1) = 1;
stBitPacking.bBit31 := (SHR(nSeed, 31) AND 1) = 1;
stBitPacking.bBit32 := (SHR(nSeed, 32) AND 1) = 1;
stBitPacking.bBit33 := (SHR(nSeed, 33) AND 1) = 1;
stBitPacking.bBit34 := (SHR(nSeed, 34) AND 1) = 1;
stBitPacking.bBit35 := (SHR(nSeed, 35) AND 1) = 1;
stBitPacking.bBit36 := (SHR(nSeed, 36) AND 1) = 1;
stBitPacking.bBit37 := (SHR(nSeed, 37) AND 1) = 1;
stBitPacking.bBit38 := (SHR(nSeed, 38) AND 1) = 1;
stBitPacking.bBit39 := (SHR(nSeed, 39) AND 1) = 1;
stBitPacking.bBit40 := (SHR(nSeed, 40) AND 1) = 1;
stBitPacking.bBit41 := (SHR(nSeed, 41) AND 1) = 1;
stBitPacking.bBit42 := (SHR(nSeed, 42) AND 1) = 1;
stBitPacking.bBit43 := (SHR(nSeed, 43) AND 1) = 1;
stBitPacking.bBit44 := (SHR(nSeed, 44) AND 1) = 1;
stBitPacking.bBit45 := (SHR(nSeed, 45) AND 1) = 1;
stBitPacking.bBit46 := (SHR(nSeed, 46) AND 1) = 1;
stBitPacking.bBit47 := (SHR(nSeed, 47) AND 1) = 1;
stBitPacking.bBit48 := (SHR(nSeed, 48) AND 1) = 1;
stBitPacking.bBit49 := (SHR(nSeed, 49) AND 1) = 1;
stBitPacking.bBit50 := (SHR(nSeed, 50) AND 1) = 1;
stBitPacking.bBit51 := (SHR(nSeed, 51) AND 1) = 1;
stBitPacking.bBit52 := (SHR(nSeed, 52) AND 1) = 1;
stBitPacking.bBit53 := (SHR(nSeed, 53) AND 1) = 1;
stBitPacking.bBit54 := (SHR(nSeed, 54) AND 1) = 1;
stBitPacking.bBit55 := (SHR(nSeed, 55) AND 1) = 1;
stBitPacking.bBit56 := (SHR(nSeed, 56) AND 1) = 1;
stBitPacking.bBit57 := (SHR(nSeed, 57) AND 1) = 1;
stBitPacking.bBit58 := (SHR(nSeed, 58) AND 1) = 1;
stBitPacking.bBit59 := (SHR(nSeed, 59) AND 1) = 1;
stBitPacking.bBit60 := (SHR(nSeed, 60) AND 1) = 1;
stBitPacking.bBit61 := (SHR(nSeed, 61) AND 1) = 1;
stBitPacking.bBit62 := (SHR(nSeed, 62) AND 1) = 1;
stBitPacking.bBit63 := (SHR(nSeed, 63) AND 1) = 1;

//FB_Init is always available implicitly and it is used primarily for initialization.
//The return value is not evaluated. For a specific influence, you can also declare the
//methods explicitly and provide additional code there with the standard initialization
//code. You can evaluate the return value.
METHOD FB_Init: BOOL
VAR_INPUT
    bInitRetains : BOOL; // TRUE: the retain variables are initialized (reset warm / reset cold)
    bInCopyCode : BOOL;  // TRUE: the instance will be copied to the copy code afterward (online change)
	nSeed : REFERENCE TO ULINT;
END_VAR
THIS^.nSeed REF= nSeed;
END_METHOD

END_FUNCTION_BLOCK

// ---- Lib/Arrays/FB_ArrayTest.TcPOU
FUNCTION_BLOCK FB_ArrayTest
VAR
	// Control
	nSeed : REFERENCE TO ULINT;

	// Scratch (derived-value working storage, not seed-test outputs)
	nSeedSt1 : ULINT;
	nScratch : ULINT;

	// Outputs
	(*
	 * Struct with an array inside -- three different array shapes as sibling
	 * members (arr1-arr3 above), not nested inside each other. This is the
	 * inverse of the "array of structs" case already covered elsewhere: here
	 * the struct-member traversal path (not the array-element path) is what
	 * has to independently reset/build each member's own arrayType tagging.
	 * If tagging leaked between siblings -- e.g. arr2's chain-boundary state
	 * bleeding into arr3's first dimension -- this is the shape that would
	 * catch it, since the three members sit directly next to each other with
	 * no array-of-array or struct-of-struct indirection to isolate them first.
	 *)
	st1 : ST_Array;
	 
	(*
	 * ARRAY-in-STRUCT-in-ARRAY: Tests whether the arrayType tag correctly
	 * resets/doesn't leak when addOffsetDepth transitions from array-element
	 * expansion into struct-member expansion — a real risk given the tag
	 * propagation is pointer-based.
	 *)
	arr1 : ARRAY[0..2,0..2] OF INT;
	 
	(*
	 * A multi-dim link immediately followed by another multi-dim link: two
	 * 2-dim links back to back (a[i,j][k,l]). More demanding than arr1 since
	 * every side of this chain boundary is multi-dim itself, not a single
	 * flat declaration with no boundary at all.
	 *)
	arr2 : ARRAY[0..1,0..1] OF ARRAY[0..1,0..1] OF INT;

	(*
	 * 3+ dims in one link, chained further: stresses that nothing hardcodes
	 * "at most 2 dims merge."
	 *)
	arr3 : ARRAY[0..1,0..1,0..1] OF ARRAY[0..1] OF INT;
	 
	(*
	 * Degenerate single-element dimension: a dimension with exactly 1 element
	 * (Elements=1), good for off-by-one bugs in the bound/overflow math.
	 *)
	arr4: ARRAY[5..5] OF ARRAY[0..9] OF INT;
	 
	(*
	 * Negative bounds on both sides of a mixed boundary: negative bounds
	 * combined with multi-dim and chaining at once (each individually tested
	 * already per the fork's history, never together).
	 *)
	arr5 : ARRAY[-5..5,-3..3] OF ARRAY[-9..-1] OF INT;
	
	(*
	 * Enum as the leaf type: does *Array.Elems end up holding Enum values
	 * correctly, and does isEnumDataType's special-casing (which already exists
	 * to stop enums being expanded as structs) interact safely with the new
	 * array-kind tagging.
	 *)
	arr6 : ARRAY[0..2,0..2] OF E_ArrayEnum;
	
	(*
	 * BIT-packed struct as the leaf type, multi-dim: combines two independent
	 * offset-math systems (bit-packing offsets, array multi-dim offsets) that
	 * have each been tested alone but maybe never together.
	 *)
	arr7 : ARRAY[0..2,0..2] OF ST_ArrayBits;
	
	(*
	 * 4+ level deep pure chain — just recursion depth, to make sure nothing
	 * assumes "at most 2 or 3 links."
	 *)
	arr8 : ARRAY[0..1] OF ARRAY[0..1] OF ARRAY[0..1] OF ARRAY[0..1] OF INT;
	
	(*
	 * 4 multi-dim links chained: Stresses both axes at once. nothing may assume
	 * "at most N links" (arr8's test) AND nothing may assume "a chain boundary
	 * only ever follows a single-dim link" (arr8's three links are all
	 * single-dim, giving it a fallback shape to lean on; this one has none)
	 * -- every one of the three chain boundaries must restart bracket
	 * nesting while two real dims merge via comma on *both* sides of it,
	 * four times over, with no single-dim link anywhere to paper over an
	 * off-by-one in "same declaration vs new declaration."
	 *)
	arr9 : ARRAY[0..1, 0..1] OF ARRAY[0..1, 0..1] OF ARRAY[0..1, 0..1] OF ARRAY[0..1, 0..1] OF INT;

	// Private
	// loop variables
	i : DINT;
	j : DINT;
	k : DINT;
	l : DINT;
	m : DINT;
	n : DINT;
	o : DINT;
	p : DINT;
END_VAR

// st1 -- offset seed, same shapes as arr1/arr2/arr3
nSeedSt1 := nSeed + 1000000;
FOR i := 0 TO 2 DO
    FOR j := 0 TO 2 DO
        st1.arr1[i,j] := DINT_TO_INT(ULINT_TO_DINT(nSeedSt1) + i*2 + j*3);
    END_FOR
END_FOR
FOR i := 0 TO 1 DO
    FOR j := 0 TO 1 DO
        FOR k := 0 TO 1 DO
            FOR l := 0 TO 1 DO
                st1.arr2[i,j][k,l] := DINT_TO_INT(ULINT_TO_DINT(nSeedSt1) + i*2 + j*3 + k*5 + l*7);
            END_FOR
        END_FOR
    END_FOR
END_FOR
FOR i := 0 TO 1 DO
    FOR j := 0 TO 1 DO
        FOR k := 0 TO 1 DO
            FOR l := 0 TO 1 DO
                st1.arr3[i,j,k][l] := DINT_TO_INT(ULINT_TO_DINT(nSeedSt1) + i*2 + j*3 + k*5 + l*7);
            END_FOR
        END_FOR
    END_FOR
END_FOR

// arr1 : ARRAY[0..2,0..2] OF INT
FOR i := 0 TO 2 DO
    FOR j := 0 TO 2 DO
        arr1[i,j] := DINT_TO_INT(ULINT_TO_DINT(nSeed) + i*2 + j*3);
    END_FOR
END_FOR

// arr2 : ARRAY[0..1,0..1] OF ARRAY[0..1,0..1] OF INT
FOR i := 0 TO 1 DO
    FOR j := 0 TO 1 DO
        FOR k := 0 TO 1 DO
            FOR l := 0 TO 1 DO
                arr2[i,j][k,l] := DINT_TO_INT(ULINT_TO_DINT(nSeed) + i*2 + j*3 + k*5 + l*7);
            END_FOR
        END_FOR
    END_FOR
END_FOR

// arr3 : ARRAY[0..1,0..1,0..1] OF ARRAY[0..1] OF INT
FOR i := 0 TO 1 DO
    FOR j := 0 TO 1 DO
        FOR k := 0 TO 1 DO
            FOR l := 0 TO 1 DO
                arr3[i,j,k][l] := DINT_TO_INT(ULINT_TO_DINT(nSeed) + i*2 + j*3 + k*5 + l*7);
            END_FOR
        END_FOR
    END_FOR
END_FOR

// arr4 : ARRAY[5..5] OF ARRAY[0..9] OF INT (degenerate outer dim)
FOR i := 5 TO 5 DO
    FOR j := 0 TO 9 DO
        arr4[i][j] := DINT_TO_INT(ULINT_TO_DINT(nSeed) + i*2 + j*3);
    END_FOR
END_FOR

// arr5 : ARRAY[-5..5,-3..3] OF ARRAY[-9..-1] OF INT (negative bounds, multi-dim + chained)
FOR i := -5 TO 5 DO
    FOR j := -3 TO 3 DO
        FOR k := -9 TO -1 DO
            arr5[i,j][k] := DINT_TO_INT(ULINT_TO_DINT(nSeed) + i*2 + j*3 + k*5);
        END_FOR
    END_FOR
END_FOR

// arr6 : ARRAY[0..2,0..2] OF E_ArrayEnum
FOR i := 0 TO 2 DO
    FOR j := 0 TO 2 DO
        nScratch := nSeed + DINT_TO_UDINT(i)*2 + DINT_TO_UDINT(j)*3;
        CASE nScratch MOD 4 OF
			1: arr6[i,j] := E_ArrayEnum.Member2;
			2: arr6[i,j] := E_ArrayEnum.Member3;
			3: arr6[i,j] := E_ArrayEnum.Member4;
		ELSE
			arr6[i,j] := E_ArrayEnum.Member1;
		END_CASE
    END_FOR
END_FOR

// arr7 : ARRAY[0..2,0..2] OF ST_ArrayBits (64-bit pattern, bulk copy)
FOR i := 0 TO 2 DO
    FOR j := 0 TO 2 DO
        nScratch := nSeed + DINT_TO_ULINT(i)*2 + DINT_TO_ULINT(j)*3;
        MEMCPY(ADR(arr7[i,j]), ADR(nScratch), SIZEOF(arr7[i,j]));
    END_FOR
END_FOR

// arr8 : 4 single-dim links chained
FOR i := 0 TO 1 DO
    FOR j := 0 TO 1 DO
        FOR k := 0 TO 1 DO
            FOR l := 0 TO 1 DO
                arr8[i][j][k][l] := DINT_TO_INT(ULINT_TO_DINT(nSeed) + i*2 + j*3 + k*5 + l*7);
            END_FOR
        END_FOR
    END_FOR
END_FOR

// arr9 : 4 chained 2-D links (8 indices)
FOR i := 0 TO 1 DO
 FOR j := 0 TO 1 DO
  FOR k := 0 TO 1 DO
   FOR l := 0 TO 1 DO
    FOR m := 0 TO 1 DO
     FOR n := 0 TO 1 DO
      FOR o := 0 TO 1 DO
       FOR p := 0 TO 1 DO
        arr9[i,j][k,l][m,n][o,p] := DINT_TO_INT(ULINT_TO_DINT(nSeed) + i*2 + j*3 + k*5 + l*7 + m*11 + n*13 + o*17 + p*19);
       END_FOR
      END_FOR
     END_FOR
    END_FOR
   END_FOR
  END_FOR
 END_FOR
END_FOR

//FB_Init is always available implicitly and it is used primarily for initialization.
//The return value is not evaluated. For a specific influence, you can also declare the
//methods explicitly and provide additional code there with the standard initialization
//code. You can evaluate the return value.
METHOD FB_Init: BOOL
VAR_INPUT
    bInitRetains : BOOL; // TRUE: the retain variables are initialized (reset warm / reset cold)
    bInCopyCode : BOOL;  // TRUE: the instance will be copied to the copy code afterward (online change)
	nSeed : REFERENCE TO ULINT;
END_VAR
THIS^.nSeed REF= nSeed;
END_METHOD

END_FUNCTION_BLOCK

// ---- Lib/Writing/FB_WriteTest.TcPOU
FUNCTION_BLOCK FB_WriteTest
VAR
	// Writable targets — PLC never modifies these, Go test owns them
	bBoolVar : BOOL;
	nSintVar : SINT;
	nUsintVar : USINT;
	nByteVar : BYTE;
	nIntVar : INT;
	nUintVar : UINT;
	nWordVar : WORD;
	nDintVar : DINT;
	nUdintVar : UDINT;
	nDwordVar : DWORD;
	nLintVar : LINT;
	nUlintVar : ULINT;
	nLwordVar : LWORD;
	fRealVar : REAL;
	fLrealVar : LREAL;
	tTimeVar : TIME;
	tdTimeOfDayVar : TOD;
	dDateVar : DATE;
	dtDateTimeVar : DT;
	tLtimeVar : LTIME;
	tdLTimeOfDayVar : LTOD;
	dLDateVar : LDATE;
	dtLDateTimeVar : LDT;
	sStringVar : STRING(255);
	stStructVar : ST_TypeTestStruct;
	aIntArray : ARRAY[0..9] OF INT;
	aDintArray : ARRAY[0..9] OF DINT;
	aIntArray2d : ARRAY[0..2, 0..2] OF INT;
END_VAR

END_FUNCTION_BLOCK

// ---- Lib/Gvl/FB_GvlTest.TcPOU
FUNCTION_BLOCK FB_GvlTest
VAR
	// Control
	nSeed : REFERENCE TO ULINT;

	// Private
	nLoopIndex1 : UDINT;
	nLoopIndex2 : UDINT;
END_VAR

// -----------------------------------------------------------------------
// Update variables — all fields are deterministic functions of seed
// -----------------------------------------------------------------------
GVL_Test.bBoolVar := (nSeed MOD 2 = 0);
GVL_Test.nSintVar := ULINT_TO_SINT(nSeed);
GVL_Test.nUsintVar := ULINT_TO_USINT(nSeed);
GVL_Test.nByteVar := ULINT_TO_BYTE(nSeed);
GVL_Test.nIntVar := ULINT_TO_INT(nSeed);
GVL_Test.nUintVar := ULINT_TO_UINT(nSeed);
GVL_Test.nWordVar := ULINT_TO_WORD(nSeed);
GVL_Test.nDintVar := ULINT_TO_DINT(nSeed);
GVL_Test.nUdintVar := ULINT_TO_UDINT(nSeed);
GVL_Test.nDwordVar := ULINT_TO_DWORD(nSeed);
GVL_Test.nLintVar := ULINT_TO_LINT(nSeed);
GVL_Test.nUlintVar := nSeed;
GVL_Test.nLwordVar := ULINT_TO_LWORD(nSeed);
GVL_Test.fRealVar := ULINT_TO_REAL(nSeed);
GVL_Test.fLrealVar := ULINT_TO_LREAL(nSeed);

// Date/time types — raw truncating casts, same bit pattern Go test will verify
GVL_Test.tTimeVar := ULINT_TO_TIME(nSeed);
GVL_Test.tdTimeOfDayVar := ULINT_TO_TOD(nSeed MOD 86400000);
GVL_Test.dDateVar := ULINT_TO_DATE(nSeed);
GVL_Test.dtDateTimeVar := ULINT_TO_DT(nSeed);
GVL_Test.tLTimeVar := ULINT_TO_LTIME(nSeed);
GVL_Test.tdLTimeOfDayVar  := ULINT_TO_LTOD(nSeed MOD 86400000000000);
GVL_Test.dLDateVar := ULINT_TO_LDATE(nSeed);
GVL_Test.dtLDateTimeVar := ULINT_TO_LDT(nSeed);
GVL_Test.sStringVar := CONCAT('S=', ULINT_TO_STRING(nSeed));

// -----------------------------------------------------------------------
// Update test struct — all fields are deterministic functions of seed
// -----------------------------------------------------------------------
GVL_Test.stStructVar.nSeed := ULINT_TO_UDINT(nSeed);
GVL_Test.stStructVar.bBoolVar := GVL_Test.bBoolVar;
GVL_Test.stStructVar.nSintVar := GVL_Test.nSintVar;
GVL_Test.stStructVar.nUsintVar := GVL_Test.nUsintVar;
GVL_Test.stStructVar.nByteVar := GVL_Test.nByteVar;
GVL_Test.stStructVar.nIntVar := GVL_Test.nIntVar;
GVL_Test.stStructVar.nUintVar := GVL_Test.nUintVar;
GVL_Test.stStructVar.nWordVar := GVL_Test.nWordVar;
GVL_Test.stStructVar.nDintVar := GVL_Test.nDintVar;
GVL_Test.stStructVar.nUdintVar := GVL_Test.nUdintVar;
GVL_Test.stStructVar.nDwordVar := GVL_Test.nDwordVar;
GVL_Test.stStructVar.nLintVar := GVL_Test.nLintVar;
GVL_Test.stStructVar.nUlintVar := GVL_Test.nUlintVar;
GVL_Test.stStructVar.nLwordVar := GVL_Test.nLwordVar;
GVL_Test.stStructVar.fRealVar := GVL_Test.fRealVar;
GVL_Test.stStructVar.fLrealVar := GVL_Test.fLrealVar;
GVL_Test.stStructVar.tTimeVar := GVL_Test.tTimeVar;
GVL_Test.stStructVar.tdTimeOfDayVar := GVL_Test.tdTimeOfDayVar;
GVL_Test.stStructVar.dDateVar := GVL_Test.dDateVar;
GVL_Test.stStructVar.dtDateTimeVar := GVL_Test.dtDateTimeVar;
GVL_Test.stStructVar.tLTimeVar := GVL_Test.tLTimeVar;
GVL_Test.stStructVar.tdLTimeOfDayVar := GVL_Test.tdLTimeOfDayVar;
GVL_Test.stStructVar.dLDateVar := GVL_Test.dLDateVar;
GVL_Test.stStructVar.dtLDateTimeVar := GVL_Test.dtLDateTimeVar;
GVL_Test.stStructVar.sStringVar := GVL_Test.sStringVar;

// -----------------------------------------------------------------------
// Update 1-D arrays: element[i] = UDINT_TO_x(seed + i)
// -----------------------------------------------------------------------
FOR nLoopIndex1 := 0 TO 9 DO
	GVL_Test.aIntArray[nLoopIndex1] := ULINT_TO_INT(nSeed + nLoopIndex1);
	GVL_Test.aDintArray[nLoopIndex1] := ULINT_TO_DINT(nSeed + nLoopIndex1);
END_FOR

// -----------------------------------------------------------------------
// Update 2-D array: element[i,j] = UDINT_TO_INT(seed + i*3 + j)
// -----------------------------------------------------------------------
FOR nLoopIndex1 := 0 TO 2 DO
	FOR nLoopIndex2 := 0 TO 2 DO
		GVL_Test.aIntArray2d[nLoopIndex1, nLoopIndex2] := ULINT_TO_INT(nSeed + nLoopIndex1 * 3 + nLoopIndex2);
	END_FOR
END_FOR

//FB_Init is always available implicitly and it is used primarily for initialization.
//The return value is not evaluated. For a specific influence, you can also declare the
//methods explicitly and provide additional code there with the standard initialization
//code. You can evaluate the return value.
METHOD FB_Init: BOOL
VAR_INPUT
    bInitRetains : BOOL; // TRUE: the retain variables are initialized (reset warm / reset cold)
    bInCopyCode : BOOL;  // TRUE: the instance will be copied to the copy code afterward (online change)
	nSeed : REFERENCE TO ULINT;
END_VAR
THIS^.nSeed REF= nSeed;
END_METHOD

END_FUNCTION_BLOCK

// ---- Lib/Attributes/FB_AttributeTest.TcPOU
{attribute 'linkalways'}
{attribute 'some_made_up_key':='some_made_up_value'}
FUNCTION_BLOCK FB_AttributeTest
VAR
END_VAR

END_FUNCTION_BLOCK
